TYPE E_LintEnum :
(
    eIdle := 0,
    eRun,
    eErr := 10
);
END_TYPE

(* stored: Version 1.1.0.1, ProductVersion 3.1.4024.16
   DUT E_LintEnum: Id {d728de05-b056-4884-8476-39202d90bd59} *)
